Staubli VAL3: do_for.pgx

public program do_for(string x_sKey, num x_nIndex)
  local num l_nIOindex
  local bool l_bResult
  local num l_nLoop
  local bool l_bErr
  local bool l_bActive
  local string l_skey
  local num l_i
  local string l_sType
begin
  waitEndMove()
  l_bActive=false
  if progTemp:pProgItem[x_sKey].pProgTemplate[x_nIndex].fForItem.sIOindex=="value"
    l_nLoop=progTemp:pProgItem[x_sKey].pProgTemplate[x_nIndex].fForItem.nLoopValue
    l_bActive=true
  else
    toNum(progTemp:pProgItem[x_sKey].pProgTemplate[x_nIndex].fForItem.sIOindex,l_nIOindex,l_bResult)
    if l_bResult
      call io:getAnaIO(io:aInItem[l_nIOindex].aAio,l_nLoop,l_bErr)
      l_bActive=true
    endIf
  endIf
  l_skey=progTemp:pProgItem[x_sKey].pProgTemplate[x_nIndex].fForItem.sForTRAJ
  l_sType=progTemp:pProgItem[x_sKey].pProgTemplate[x_nIndex].sTRAJname
  switch l_sType
    case "PROG"
      if l_bActive
        for l_i = 0 to l_nLoop
          call makeTraj(l_skey)
        endFor
      endIf
    break
    case "TRAJ"
      if l_bActive
        for l_i = 0 to l_nLoop
          call trajectory:makeTraj(l_skey)
        endFor
      endIf
    break
  endSwitch

end
